(* IEC 61131-3 sources: Pirate/PLC/POU, 5 files *)

(* ---- EcrireSorties.st ---- *)
FUNCTION EcrireSorties : BOOL
// POU autonome extrait de FB_InterfacePIRATE (branche dev).
// A appeler APRES le calcul du simulateur.
// Reproduit uniquement les copies de variables GVL ; aucun mapping BFS ajoute.
// Appeler apres la simulation.
GVL_PIRATE.ST_THEGONNEC_AT2_Defaut_Auto_transfo_2 := GVL_PIRATE_Interne.S_ST_THEGONNEC_AT2_Defaut_Auto_transfo_2;
GVL_PIRATE.ST_THEGONNEC_SYSTEME_PC_SNCF_PA_Defaut_Controle_General := GVL_PIRATE_Interne.S_ST_THEGONNEC_SYSTEME_PC_SNCF_PA_Defaut_Controle_General;
GVL_PIRATE.ST_THEGONNEC_U_Cat__TT_2C_Etat_tension_voie_2 := GVL_PIRATE_Interne.S_ST_THEGONNEC_U_Cat__TT_2C_Etat_tension_voie_2;
GVL_PIRATE.ST_THEGONNEC_U_Cat__TT_3C_Etat_tension_voie_1 := GVL_PIRATE_Interne.S_ST_THEGONNEC_U_Cat__TT_3C_Etat_tension_voie_1;
GVL_PIRATE.ST_THEGONNEC_AT1_Defaut_Auto_transfo_1 := GVL_PIRATE_Interne.S_ST_THEGONNEC_AT1_Defaut_Auto_transfo_1;
GVL_PIRATE.BREST_SYSTEME_PC_SNCF_PA_Defaut_Controle_General := GVL_PIRATE_Interne.S_BREST_SYSTEME_PC_SNCF_PA_Defaut_Controle_General;
GVL_PIRATE.BREST_SA_Defaut_Chauffage_Commandes := GVL_PIRATE_Interne.S_BREST_SA_Defaut_Chauffage_Commandes;
GVL_PIRATE.BREST_U_Cat__TT_IA6_Etat_tension_voie := GVL_PIRATE_Interne.S_BREST_U_Cat__TT_IA6_Etat_tension_voie;
GVL_PIRATE.BREST_U_Cat__TT_IA1_Etat_tension_voie := GVL_PIRATE_Interne.S_BREST_U_Cat__TT_IA1_Etat_tension_voie;
GVL_PIRATE.BREST_U_Cat__TT_2C_Etat_tension_voie_2 := GVL_PIRATE_Interne.S_BREST_U_Cat__TT_2C_Etat_tension_voie_2;
GVL_PIRATE.PENCRAN_1_U_Feeder_TT_3F_Etat_tension_voie_1 := GVL_PIRATE_Interne.S_PENCRAN_1_U_Feeder_TT_3F_Etat_tension_voie_1;
GVL_PIRATE.PENCRAN_1_U_Feeder_TT_4F_Etat_tension_voie_2 := GVL_PIRATE_Interne.S_PENCRAN_1_U_Feeder_TT_4F_Etat_tension_voie_2;
GVL_PIRATE.PENCRAN_1_TT_Feeder_DL_Etat_tension := GVL_PIRATE_Interne.S_PENCRAN_1_TT_Feeder_DL_Etat_tension;
GVL_PIRATE.PENCRAN_1_U_Cat__TT_2C_Etat_tension_voie_2 := GVL_PIRATE_Interne.S_PENCRAN_1_U_Cat__TT_2C_Etat_tension_voie_2;
GVL_PIRATE.PENCRAN_1_U_Cat__TT_4C_Etat_tension_voie_2 := GVL_PIRATE_Interne.S_PENCRAN_1_U_Cat__TT_4C_Etat_tension_voie_2;
GVL_PIRATE.PENCRAN_1_U_Feeder_TT_1F_Etat_tension_voie_1 := GVL_PIRATE_Interne.S_PENCRAN_1_U_Feeder_TT_1F_Etat_tension_voie_1;
GVL_PIRATE.PENCRAN_1_U_Cat__TT_3C_Etat_tension_voie_1 := GVL_PIRATE_Interne.S_PENCRAN_1_U_Cat__TT_3C_Etat_tension_voie_1;
GVL_PIRATE.PENCRAN_1_U_Cat__TT_1C_Etat_tension_voie_1 := GVL_PIRATE_Interne.S_PENCRAN_1_U_Cat__TT_1C_Etat_tension_voie_1;
GVL_PIRATE.PENCRAN_1_TT_Cat__DB_Etat_tension := GVL_PIRATE_Interne.S_PENCRAN_1_TT_Cat__DB_Etat_tension;
GVL_PIRATE.PENCRAN_1_U_Feeder_TT_2F_Etat_tension_voie_2 := GVL_PIRATE_Interne.S_PENCRAN_1_U_Feeder_TT_2F_Etat_tension_voie_2;
GVL_PIRATE.PENCRAN_1_SYSTEME_PC_SNCF_PA_Defaut_Controle_General := GVL_PIRATE_Interne.S_PENCRAN_1_SYSTEME_PC_SNCF_PA_Defaut_Controle_General;
GVL_PIRATE.PENCRAN_1_TT_Cat__DL_Etat_tension := GVL_PIRATE_Interne.S_PENCRAN_1_TT_Cat__DL_Etat_tension;
GVL_PIRATE.PENCRAN_1_TT_Feeder_DB_Etat_tension := GVL_PIRATE_Interne.S_PENCRAN_1_TT_Feeder_DB_Etat_tension;
GVL_PIRATE.PENCRAN_1_GT2_Defaut_Alim__Protection__W_D_ := GVL_PIRATE_Interne.S_PENCRAN_1_GT2_Defaut_Alim__Protection__W_D_;
GVL_PIRATE.PENCRAN_1_DL__TSS__Defaut_Alim__Protection__W_D_ := GVL_PIRATE_Interne.S_PENCRAN_1_DL__TSS__Defaut_Alim__Protection__W_D_;
GVL_PIRATE.PENCRAN_1_GT1_Defaut_Alim__Protection__W_D_ := GVL_PIRATE_Interne.S_PENCRAN_1_GT1_Defaut_Alim__Protection__W_D_;
GVL_PIRATE.PENCRAN_1_GT1_Defaut_Transfo__Groupe_Traction := GVL_PIRATE_Interne.S_PENCRAN_1_GT1_Defaut_Transfo__Groupe_Traction;
GVL_PIRATE.PENCRAN_1_GT2_Defaut_Transfo__Groupe_Traction := GVL_PIRATE_Interne.S_PENCRAN_1_GT2_Defaut_Transfo__Groupe_Traction;
GVL_PIRATE.PENCRAN_1_DL__TSS__Defaut_SF6 := GVL_PIRATE_Interne.S_PENCRAN_1_DL__TSS__Defaut_SF6;
GVL_PIRATE.PENCRAN_1_SA_Defaut_Chargeur := GVL_PIRATE_Interne.S_PENCRAN_1_SA_Defaut_Chargeur;
GVL_PIRATE.PENCRAN_1_D2___25kV_Defaut_SF6_2eme_seuil := GVL_PIRATE_Interne.S_PENCRAN_1_D2___25kV_Defaut_SF6_2eme_seuil;
GVL_PIRATE.PENCRAN_1_DB__TSS__Defaut_Alim__Protection__W_D_ := GVL_PIRATE_Interne.S_PENCRAN_1_DB__TSS__Defaut_Alim__Protection__W_D_;
GVL_PIRATE.PENCRAN_1_Automate_Defaut_Relais_PROM := GVL_PIRATE_Interne.S_PENCRAN_1_Automate_Defaut_Relais_PROM;
GVL_PIRATE.PENCRAN_1_D2___25kV_Defaut_Commande_disjoncteur := GVL_PIRATE_Interne.S_PENCRAN_1_D2___25kV_Defaut_Commande_disjoncteur;
GVL_PIRATE.PENCRAN_1_Automate_Defaut_Reenclencheur := GVL_PIRATE_Interne.S_PENCRAN_1_Automate_Defaut_Reenclencheur;
GVL_PIRATE.PENCRAN_1_DB__TSS__Defaut_SF6 := GVL_PIRATE_Interne.S_PENCRAN_1_DB__TSS__Defaut_SF6;
GVL_PIRATE.LANDIVISIAU_AT2_Defaut_Auto_transfo_2 := GVL_PIRATE_Interne.S_LANDIVISIAU_AT2_Defaut_Auto_transfo_2;
GVL_PIRATE.LANDIVISIAU_U_Cat__TT_2C_Etat_tension_voie_2 := GVL_PIRATE_Interne.S_LANDIVISIAU_U_Cat__TT_2C_Etat_tension_voie_2;
GVL_PIRATE.LANDIVISIAU_AT1_Defaut_Auto_transfo_1 := GVL_PIRATE_Interne.S_LANDIVISIAU_AT1_Defaut_Auto_transfo_1;
GVL_PIRATE.LANDIVISIAU_SYSTEME_PC_SNCF_PA_Defaut_Controle_General := GVL_PIRATE_Interne.S_LANDIVISIAU_SYSTEME_PC_SNCF_PA_Defaut_Controle_General;
GVL_PIRATE.LANDIVISIAU_U_Cat__TT_3C_Etat_tension_voie_1 := GVL_PIRATE_Interne.S_LANDIVISIAU_U_Cat__TT_3C_Etat_tension_voie_1;
GVL_PIRATE.ST_MARC_U_Cat__TT_3C_Etat_tension_voie_1 := GVL_PIRATE_Interne.S_ST_MARC_U_Cat__TT_3C_Etat_tension_voie_1;
GVL_PIRATE.ST_MARC_SYSTEME_PC_SNCF_PA_Defaut_Controle_General := GVL_PIRATE_Interne.S_ST_MARC_SYSTEME_PC_SNCF_PA_Defaut_Controle_General;
GVL_PIRATE.ST_MARC_AT1_Defaut_Auto_transfo_1 := GVL_PIRATE_Interne.S_ST_MARC_AT1_Defaut_Auto_transfo_1;
GVL_PIRATE.ST_MARC_U_Cat__TT_2C_Etat_tension_voie_2 := GVL_PIRATE_Interne.S_ST_MARC_U_Cat__TT_2C_Etat_tension_voie_2;
GVL_PIRATE.ST_MARC_AT2_Defaut_Auto_transfo_2 := GVL_PIRATE_Interne.S_ST_MARC_AT2_Defaut_Auto_transfo_2;
GVL_PIRATE.LA_FOREST_AT_Defaut_Auto_transfo := GVL_PIRATE_Interne.S_LA_FOREST_AT_Defaut_Auto_transfo;
GVL_PIRATE.LA_FOREST_SYSTEME_PC_SNCF_PA_Defaut_Controle_General := GVL_PIRATE_Interne.S_LA_FOREST_SYSTEME_PC_SNCF_PA_Defaut_Controle_General;
GVL_PIRATE.KERIVIN_SYSTEME_PC_SNCF_PA_Defaut_Controle_General := GVL_PIRATE_Interne.S_KERIVIN_SYSTEME_PC_SNCF_PA_Defaut_Controle_General;
GVL_PIRATE.KERIVIN_U_Cat__TT_2C_Etat_tension_voie_2 := GVL_PIRATE_Interne.S_KERIVIN_U_Cat__TT_2C_Etat_tension_voie_2;
GVL_PIRATE.KERIVIN_AT2_Defaut_Auto_transfo_2 := GVL_PIRATE_Interne.S_KERIVIN_AT2_Defaut_Auto_transfo_2;
GVL_PIRATE.KERIVIN_AT1_Defaut_Auto_transfo_1 := GVL_PIRATE_Interne.S_KERIVIN_AT1_Defaut_Auto_transfo_1;
GVL_PIRATE.KERIVIN_U_Cat__TT_3C_Etat_tension_voie_1 := GVL_PIRATE_Interne.S_KERIVIN_U_Cat__TT_3C_Etat_tension_voie_1;
GVL_PIRATE.LANDERNEAU_SYSTEME_PC_SNCF_PA_Defaut_Controle_General := GVL_PIRATE_Interne.S_LANDERNEAU_SYSTEME_PC_SNCF_PA_Defaut_Controle_General;
GVL_PIRATE.MORLAIX_SYSTEME_PC_SNCF_PA_Defaut_Controle_General := GVL_PIRATE_Interne.S_MORLAIX_SYSTEME_PC_SNCF_PA_Defaut_Controle_General;
GVL_PIRATE.PLOUIGNEAU_U_Cat__TT_3C_Etat_tension_voie_1 := GVL_PIRATE_Interne.S_PLOUIGNEAU_U_Cat__TT_3C_Etat_tension_voie_1;
GVL_PIRATE.PLOUIGNEAU_U_Cat__TT_2C_Etat_tension_voie_2 := GVL_PIRATE_Interne.S_PLOUIGNEAU_U_Cat__TT_2C_Etat_tension_voie_2;
GVL_PIRATE.PLOUIGNEAU_AT1_Defaut_Auto_transfo_1 := GVL_PIRATE_Interne.S_PLOUIGNEAU_AT1_Defaut_Auto_transfo_1;
GVL_PIRATE.PLOUIGNEAU_U_Cat__TT_4C_Etat_tension_voie_2 := GVL_PIRATE_Interne.S_PLOUIGNEAU_U_Cat__TT_4C_Etat_tension_voie_2;
GVL_PIRATE.PLOUIGNEAU_AT2_Defaut_Auto_transfo_2 := GVL_PIRATE_Interne.S_PLOUIGNEAU_AT2_Defaut_Auto_transfo_2;
GVL_PIRATE.PLOUIGNEAU_SYSTEME_PC_SNCF_PA_Defaut_Controle_General := GVL_PIRATE_Interne.S_PLOUIGNEAU_SYSTEME_PC_SNCF_PA_Defaut_Controle_General;
GVL_PIRATE.PLOUNERIN_AT2_Defaut_Auto_transfo_2 := GVL_PIRATE_Interne.S_PLOUNERIN_AT2_Defaut_Auto_transfo_2;
GVL_PIRATE.PLOUNERIN_U_Cat__TT_3C_Etat_tension_voie_1 := GVL_PIRATE_Interne.S_PLOUNERIN_U_Cat__TT_3C_Etat_tension_voie_1;
EcrireSorties := TRUE;
END_FUNCTION

(* ---- LireEntrees.st ---- *)
FUNCTION LireEntrees : BOOL
// POU autonome extrait de FB_InterfacePIRATE (branche dev).
// A appeler AVANT le calcul du simulateur.
// Reproduit uniquement les copies de variables GVL ; aucun mapping BFS ajoute.
// Appeler avant la simulation.
GVL_PIRATE_Interne.E_ST_THEGONNEC_S20_30_Sect__de_pontage_V2 := GVL_PIRATE.ST_THEGONNEC_S20_30_Sect__de_pontage_V2;
GVL_PIRATE_Interne.E_ST_THEGONNEC_SYSTEME_PC_SNCF_PA_Douteux_vu_du_PC := GVL_PIRATE.ST_THEGONNEC_SYSTEME_PC_SNCF_PA_Douteux_vu_du_PC;
GVL_PIRATE_Interne.E_ST_THEGONNEC_IL2_Inter__de_ligne_2x25kv_V2 := GVL_PIRATE.ST_THEGONNEC_IL2_Inter__de_ligne_2x25kv_V2;
GVL_PIRATE_Interne.E_ST_THEGONNEC_IL4_Inter__de_ligne_2x25kv_V2 := GVL_PIRATE.ST_THEGONNEC_IL4_Inter__de_ligne_2x25kv_V2;
GVL_PIRATE_Interne.E_ST_THEGONNEC_SAT1___25kV_Sect__alimentation_auto_transfo1 := GVL_PIRATE.ST_THEGONNEC_SAT1___25kV_Sect__alimentation_auto_transfo1;
GVL_PIRATE_Interne.E_ST_THEGONNEC_SYSTEME_PC_SNCF_PA_Titulaire := GVL_PIRATE.ST_THEGONNEC_SYSTEME_PC_SNCF_PA_Titulaire;
GVL_PIRATE_Interne.E_ST_THEGONNEC_S21_31_Sect__de_pontage_V1 := GVL_PIRATE.ST_THEGONNEC_S21_31_Sect__de_pontage_V1;
GVL_PIRATE_Interne.E_ST_THEGONNEC_SYSTEME_PA_SNCF_PA_Perte_Date := GVL_PIRATE.ST_THEGONNEC_SYSTEME_PA_SNCF_PA_Perte_Date;
GVL_PIRATE_Interne.E_ST_THEGONNEC_IL3_Inter__de_ligne_2x25kv_V1 := GVL_PIRATE.ST_THEGONNEC_IL3_Inter__de_ligne_2x25kv_V1;
GVL_PIRATE_Interne.E_ST_THEGONNEC_SA_Manque_SA := GVL_PIRATE.ST_THEGONNEC_SA_Manque_SA;
GVL_PIRATE_Interne.E_ST_THEGONNEC_SYSTEME_PA_SNCF_PA_Carte_s__TS := GVL_PIRATE.ST_THEGONNEC_SYSTEME_PA_SNCF_PA_Carte_s__TS;
GVL_PIRATE_Interne.E_ST_THEGONNEC_IMP___25kV_Interrupteur_mise_en_parallele := GVL_PIRATE.ST_THEGONNEC_IMP___25kV_Interrupteur_mise_en_parallele;
GVL_PIRATE_Interne.E_ST_THEGONNEC_IL1_Inter__de_ligne_2x25kv_V1 := GVL_PIRATE.ST_THEGONNEC_IL1_Inter__de_ligne_2x25kv_V1;
GVL_PIRATE_Interne.E_ST_THEGONNEC_SYSTEME_PC_SNCF_PA_Liaison_PC______PA := GVL_PIRATE.ST_THEGONNEC_SYSTEME_PC_SNCF_PA_Liaison_PC______PA;
GVL_PIRATE_Interne.E_ST_THEGONNEC_SYSTEME_PC_SNCF_PA_Non_date := GVL_PIRATE.ST_THEGONNEC_SYSTEME_PC_SNCF_PA_Non_date;
GVL_PIRATE_Interne.E_ST_THEGONNEC_Contrile_Local_Commande_locale_individuelle := GVL_PIRATE.ST_THEGONNEC_Contrile_Local_Commande_locale_individuelle;
GVL_PIRATE_Interne.E_ST_THEGONNEC_FICTIF_Organe_Fictif := GVL_PIRATE.ST_THEGONNEC_FICTIF_Organe_Fictif;
GVL_PIRATE_Interne.E_ST_THEGONNEC_SAT2___25kV_Sect__alimentation_auto_transfo2 := GVL_PIRATE.ST_THEGONNEC_SAT2___25kV_Sect__alimentation_auto_transfo2;
GVL_PIRATE_Interne.E_ST_THEGONNEC_SYSTEME_PA_SNCF_PA_Perte_Information := GVL_PIRATE.ST_THEGONNEC_SYSTEME_PA_SNCF_PA_Perte_Information;
GVL_PIRATE_Interne.E_ST_THEGONNEC_SYSTEME_PA_SNCF_PA_Carte_s__TC := GVL_PIRATE.ST_THEGONNEC_SYSTEME_PA_SNCF_PA_Carte_s__TC;
GVL_PIRATE_Interne.E_BREST_SA_Manque_SA := GVL_PIRATE.BREST_SA_Manque_SA;
GVL_PIRATE_Interne.E_BREST_SYSTEME_PA_SNCF_PA_Carte_s__TS := GVL_PIRATE.BREST_SYSTEME_PA_SNCF_PA_Carte_s__TS;
GVL_PIRATE_Interne.E_BREST_Contrile_Local_Commande_locale_individuelle := GVL_PIRATE.BREST_Contrile_Local_Commande_locale_individuelle;
GVL_PIRATE_Interne.E_BREST_SYSTEME_PC_SNCF_PA_Non_date := GVL_PIRATE.BREST_SYSTEME_PC_SNCF_PA_Non_date;
GVL_PIRATE_Interne.E_BREST_SYSTEME_PA_SNCF_PA_Perte_Date := GVL_PIRATE.BREST_SYSTEME_PA_SNCF_PA_Perte_Date;
GVL_PIRATE_Interne.E_BREST_SYSTEME_PC_SNCF_PA_Liaison_PC______PA := GVL_PIRATE.BREST_SYSTEME_PC_SNCF_PA_Liaison_PC______PA;
GVL_PIRATE_Interne.E_BREST_SYSTEME_PA_SNCF_PA_Perte_Information := GVL_PIRATE.BREST_SYSTEME_PA_SNCF_PA_Perte_Information;
GVL_PIRATE_Interne.E_BREST_SYSTEME_PC_SNCF_PA_Titulaire := GVL_PIRATE.BREST_SYSTEME_PC_SNCF_PA_Titulaire;
GVL_PIRATE_Interne.E_BREST_IA6_Automatisme_Automat_Ouv_PLUS_Bloc_Debloc_IA__Ouv_ := GVL_PIRATE.BREST_IA6_Automatisme_Automat_Ouv_PLUS_Bloc_Debloc_IA__Ouv_;
GVL_PIRATE_Interne.E_BREST_IL2_Inter__de_ligne_25kv_V2 := GVL_PIRATE.BREST_IL2_Inter__de_ligne_25kv_V2;
GVL_PIRATE_Interne.E_BREST_IA1_Automatisme_Automat_Ouv_PLUS_Bloc_Debloc_IA__Ouv_ := GVL_PIRATE.BREST_IA1_Automatisme_Automat_Ouv_PLUS_Bloc_Debloc_IA__Ouv_;
GVL_PIRATE_Interne.E_BREST_IA6_Interrupteur_d_Alimentation__IA_ := GVL_PIRATE.BREST_IA6_Interrupteur_d_Alimentation__IA_;
GVL_PIRATE_Interne.E_BREST_IL1_Inter__de_ligne_25kv_V1 := GVL_PIRATE.BREST_IL1_Inter__de_ligne_25kv_V1;
GVL_PIRATE_Interne.E_BREST_SYSTEME_PC_SNCF_PA_Douteux_vu_du_PC := GVL_PIRATE.BREST_SYSTEME_PC_SNCF_PA_Douteux_vu_du_PC;
GVL_PIRATE_Interne.E_BREST_IA1_Interrupteur_d_Alimentation__IA_ := GVL_PIRATE.BREST_IA1_Interrupteur_d_Alimentation__IA_;
GVL_PIRATE_Interne.E_BREST_SYSTEME_PA_SNCF_PA_Carte_s__TC := GVL_PIRATE.BREST_SYSTEME_PA_SNCF_PA_Carte_s__TC;
GVL_PIRATE_Interne.E_BREST_FICTIF_Organe_Fictif := GVL_PIRATE.BREST_FICTIF_Organe_Fictif;
GVL_PIRATE_Interne.E_PENCRAN_1_SYSTEME_PC_SNCF_PA_Douteux_vu_du_PC := GVL_PIRATE.PENCRAN_1_SYSTEME_PC_SNCF_PA_Douteux_vu_du_PC;
GVL_PIRATE_Interne.E_PENCRAN_1_SYSTEME_PA_SNCF_PA_Perte_Date := GVL_PIRATE.PENCRAN_1_SYSTEME_PA_SNCF_PA_Perte_Date;
GVL_PIRATE_Interne.E_PENCRAN_1_SYSTEME_PC_SNCF_PA_Non_date := GVL_PIRATE.PENCRAN_1_SYSTEME_PC_SNCF_PA_Non_date;
GVL_PIRATE_Interne.E_PENCRAN_1_UHT_1_Absence_tension_ligne_HT := GVL_PIRATE.PENCRAN_1_UHT_1_Absence_tension_ligne_HT;
GVL_PIRATE_Interne.E_PENCRAN_1_SYSTEME_PC_SNCF_PA_Liaison_PC______PA := GVL_PIRATE.PENCRAN_1_SYSTEME_PC_SNCF_PA_Liaison_PC______PA;
GVL_PIRATE_Interne.E_PENCRAN_1_SYSTEME_PA_SNCF_PA_Perte_Information := GVL_PIRATE.PENCRAN_1_SYSTEME_PA_SNCF_PA_Perte_Information;
GVL_PIRATE_Interne.E_PENCRAN_1_UHT_1_Fusion_fusible_s_ := GVL_PIRATE.PENCRAN_1_UHT_1_Fusion_fusible_s_;
GVL_PIRATE_Interne.E_PENCRAN_1_SYSTEME_PC_SNCF_PA_Titulaire := GVL_PIRATE.PENCRAN_1_SYSTEME_PC_SNCF_PA_Titulaire;
GVL_PIRATE_Interne.E_PENCRAN_1_UHT_2_Absence_tension_ligne_HT := GVL_PIRATE.PENCRAN_1_UHT_2_Absence_tension_ligne_HT;
GVL_PIRATE_Interne.E_PENCRAN_1_UHT_2_Fusion_fusible_s_ := GVL_PIRATE.PENCRAN_1_UHT_2_Fusion_fusible_s_;
GVL_PIRATE_Interne.E_PENCRAN_1_SLB1_Sect__de_barre_de_ligne_25Kv := GVL_PIRATE.PENCRAN_1_SLB1_Sect__de_barre_de_ligne_25Kv;
GVL_PIRATE_Interne.E_PENCRAN_1_DL_Disj_depart_2x25kV_Le_Mans := GVL_PIRATE.PENCRAN_1_DL_Disj_depart_2x25kV_Le_Mans;
GVL_PIRATE_Interne.E_PENCRAN_1_S11___63kV_Sect__de_ligne_Haute_Tension := GVL_PIRATE.PENCRAN_1_S11___63kV_Sect__de_ligne_Haute_Tension;
GVL_PIRATE_Interne.E_PENCRAN_1_SA_Manque_SA2 := GVL_PIRATE.PENCRAN_1_SA_Manque_SA2;
GVL_PIRATE_Interne.E_PENCRAN_1_IS1_Inter__de_S_Station_2x25Kv_V1 := GVL_PIRATE.PENCRAN_1_IS1_Inter__de_S_Station_2x25Kv_V1;
GVL_PIRATE_Interne.E_PENCRAN_1_SRB1___25kV_Sect__a_rupture_brusque_GT1 := GVL_PIRATE.PENCRAN_1_SRB1___25kV_Sect__a_rupture_brusque_GT1;
GVL_PIRATE_Interne.E_PENCRAN_1_SYSTEME_PA_SNCF_PA_Carte_s__TS := GVL_PIRATE.PENCRAN_1_SYSTEME_PA_SNCF_PA_Carte_s__TS;
GVL_PIRATE_Interne.E_PENCRAN_1_SA_Manque_SA1 := GVL_PIRATE.PENCRAN_1_SA_Manque_SA1;
GVL_PIRATE_Interne.E_PENCRAN_1_SA_Manque_48V_ := GVL_PIRATE.PENCRAN_1_SA_Manque_48V_;
GVL_PIRATE_Interne.E_PENCRAN_1_SYSTEME_PA_SNCF_PA_Carte_s__TC := GVL_PIRATE.PENCRAN_1_SYSTEME_PA_SNCF_PA_Carte_s__TC;
GVL_PIRATE_Interne.E_PENCRAN_1_P1_Sect__de_pontage_V1 := GVL_PIRATE.PENCRAN_1_P1_Sect__de_pontage_V1;
GVL_PIRATE_Interne.E_PENCRAN_1_SB1___25kV_Sect__de_section_de_barre_25Kv := GVL_PIRATE.PENCRAN_1_SB1___25kV_Sect__de_section_de_barre_25Kv;
GVL_PIRATE_Interne.E_PENCRAN_1_SBP1___63kV_Sect__de_section_de_barre_HT := GVL_PIRATE.PENCRAN_1_SBP1___63kV_Sect__de_section_de_barre_HT;
GVL_PIRATE_Interne.E_PENCRAN_1_IS3_Inter__de_S_Station_25Kv_V1 := GVL_PIRATE.PENCRAN_1_IS3_Inter__de_S_Station_25Kv_V1;
GVL_PIRATE_Interne.E_PENCRAN_1_P2_Sect__de_pontage_V2 := GVL_PIRATE.PENCRAN_1_P2_Sect__de_pontage_V2;
GVL_PIRATE_Interne.E_PENCRAN_1_IS2_Inter__de_S_Station_2x25Kv_V2 := GVL_PIRATE.PENCRAN_1_IS2_Inter__de_S_Station_2x25Kv_V2;
GVL_PIRATE_Interne.E_PENCRAN_1_S21___63kV_Sect__de_ligne_Haute_Tension := GVL_PIRATE.PENCRAN_1_S21___63kV_Sect__de_ligne_Haute_Tension;
GVL_PIRATE_Interne.E_PENCRAN_1_IS4_Inter__de_S_Station_2x25Kv_V2 := GVL_PIRATE.PENCRAN_1_IS4_Inter__de_S_Station_2x25Kv_V2;
GVL_PIRATE_Interne.E_PENCRAN_1_SRB2___25kV_Sect__a_rupture_brusque_GT2 := GVL_PIRATE.PENCRAN_1_SRB2___25kV_Sect__a_rupture_brusque_GT2;
GVL_PIRATE_Interne.E_PENCRAN_1_D2___63kV_Disjoncteur_Groupe_Traction_2 := GVL_PIRATE.PENCRAN_1_D2___63kV_Disjoncteur_Groupe_Traction_2;
GVL_PIRATE_Interne.E_PENCRAN_1_DB_Disj_depart_2x25kV_Brest := GVL_PIRATE.PENCRAN_1_DB_Disj_depart_2x25kV_Brest;
GVL_PIRATE_Interne.E_PENCRAN_1_D2___25kV_Alarme_SF6_1er_seuil := GVL_PIRATE.PENCRAN_1_D2___25kV_Alarme_SF6_1er_seuil;
GVL_PIRATE_Interne.E_PENCRAN_1_Automate_Relais_PROM__TC_ := GVL_PIRATE.PENCRAN_1_Automate_Relais_PROM__TC_;
GVL_PIRATE_Interne.E_PENCRAN_1_Contrile_Local_Commande_Locale := GVL_PIRATE.PENCRAN_1_Contrile_Local_Commande_Locale;
GVL_PIRATE_Interne.E_PENCRAN_1_D1___63kV_Disjoncteur_Groupe_Traction_1 := GVL_PIRATE.PENCRAN_1_D1___63kV_Disjoncteur_Groupe_Traction_1;
GVL_PIRATE_Interne.E_PENCRAN_1_VF_Veille_Franchissement__TC_ := GVL_PIRATE.PENCRAN_1_VF_Veille_Franchissement__TC_;
GVL_PIRATE_Interne.E_PENCRAN_1_FICTIF_Organe_Fictif := GVL_PIRATE.PENCRAN_1_FICTIF_Organe_Fictif;
GVL_PIRATE_Interne.E_PENCRAN_1_D2___25kV_Disjoncteur_Groupe_Traction_2 := GVL_PIRATE.PENCRAN_1_D2___25kV_Disjoncteur_Groupe_Traction_2;
GVL_PIRATE_Interne.E_LANDIVISIAU_SYSTEME_PA_SNCF_PA_Perte_Date := GVL_PIRATE.LANDIVISIAU_SYSTEME_PA_SNCF_PA_Perte_Date;
GVL_PIRATE_Interne.E_LANDIVISIAU_S30_40_Sect__de_pontage_V2 := GVL_PIRATE.LANDIVISIAU_S30_40_Sect__de_pontage_V2;
GVL_PIRATE_Interne.E_LANDIVISIAU_SYSTEME_PC_SNCF_PA_Non_date := GVL_PIRATE.LANDIVISIAU_SYSTEME_PC_SNCF_PA_Non_date;
GVL_PIRATE_Interne.E_LANDIVISIAU_S31_41_Sect__de_pontage_V1 := GVL_PIRATE.LANDIVISIAU_S31_41_Sect__de_pontage_V1;
GVL_PIRATE_Interne.E_LANDIVISIAU_IL1_Inter__de_ligne_2x25kv_V1 := GVL_PIRATE.LANDIVISIAU_IL1_Inter__de_ligne_2x25kv_V1;
GVL_PIRATE_Interne.E_LANDIVISIAU_SYSTEME_PC_SNCF_PA_Douteux_vu_du_PC := GVL_PIRATE.LANDIVISIAU_SYSTEME_PC_SNCF_PA_Douteux_vu_du_PC;
GVL_PIRATE_Interne.E_LANDIVISIAU_SYSTEME_PA_SNCF_PA_Carte_s__TS := GVL_PIRATE.LANDIVISIAU_SYSTEME_PA_SNCF_PA_Carte_s__TS;
GVL_PIRATE_Interne.E_LANDIVISIAU_IL3_Inter__de_ligne_2x25kv_V1 := GVL_PIRATE.LANDIVISIAU_IL3_Inter__de_ligne_2x25kv_V1;
GVL_PIRATE_Interne.E_LANDIVISIAU_SA_Manque_SA := GVL_PIRATE.LANDIVISIAU_SA_Manque_SA;
GVL_PIRATE_Interne.E_LANDIVISIAU_SYSTEME_PC_SNCF_PA_Liaison_PC______PA := GVL_PIRATE.LANDIVISIAU_SYSTEME_PC_SNCF_PA_Liaison_PC______PA;
GVL_PIRATE_Interne.E_LANDIVISIAU_IL2_Inter__de_ligne_2x25kv_V2 := GVL_PIRATE.LANDIVISIAU_IL2_Inter__de_ligne_2x25kv_V2;
GVL_PIRATE_Interne.E_LANDIVISIAU_IMP___25kV_Interrupteur_mise_en_parallele := GVL_PIRATE.LANDIVISIAU_IMP___25kV_Interrupteur_mise_en_parallele;
GVL_PIRATE_Interne.E_LANDIVISIAU_SAT1___25kV_Sect__alimentation_auto_transfo1 := GVL_PIRATE.LANDIVISIAU_SAT1___25kV_Sect__alimentation_auto_transfo1;
GVL_PIRATE_Interne.E_LANDIVISIAU_SYSTEME_PC_SNCF_PA_Titulaire := GVL_PIRATE.LANDIVISIAU_SYSTEME_PC_SNCF_PA_Titulaire;
GVL_PIRATE_Interne.E_LANDIVISIAU_IL4_Inter__de_ligne_2x25kv_V2 := GVL_PIRATE.LANDIVISIAU_IL4_Inter__de_ligne_2x25kv_V2;
GVL_PIRATE_Interne.E_LANDIVISIAU_SYSTEME_PA_SNCF_PA_Perte_Information := GVL_PIRATE.LANDIVISIAU_SYSTEME_PA_SNCF_PA_Perte_Information;
GVL_PIRATE_Interne.E_LANDIVISIAU_SYSTEME_PA_SNCF_PA_Carte_s__TC := GVL_PIRATE.LANDIVISIAU_SYSTEME_PA_SNCF_PA_Carte_s__TC;
GVL_PIRATE_Interne.E_LANDIVISIAU_Contrile_Local_Commande_locale_individuelle := GVL_PIRATE.LANDIVISIAU_Contrile_Local_Commande_locale_individuelle;
GVL_PIRATE_Interne.E_LANDIVISIAU_SAT2___25kV_Sect__alimentation_auto_transfo2 := GVL_PIRATE.LANDIVISIAU_SAT2___25kV_Sect__alimentation_auto_transfo2;
GVL_PIRATE_Interne.E_LANDIVISIAU_FICTIF_Organe_Fictif := GVL_PIRATE.LANDIVISIAU_FICTIF_Organe_Fictif;
GVL_PIRATE_Interne.E_ST_MARC_S4_10_Sect__de_pontage_V2 := GVL_PIRATE.ST_MARC_S4_10_Sect__de_pontage_V2;
GVL_PIRATE_Interne.E_ST_MARC_SYSTEME_PA_SNCF_PA_Perte_Information := GVL_PIRATE.ST_MARC_SYSTEME_PA_SNCF_PA_Perte_Information;
GVL_PIRATE_Interne.E_ST_MARC_IA3_Interrupteur_d_Alimentation__IA_ := GVL_PIRATE.ST_MARC_IA3_Interrupteur_d_Alimentation__IA_;
GVL_PIRATE_Interne.E_ST_MARC_SA_Manque_SA_Satellite_2 := GVL_PIRATE.ST_MARC_SA_Manque_SA_Satellite_2;
GVL_PIRATE_Interne.E_ST_MARC_IL2_Inter__de_ligne_2x25kv_V2 := GVL_PIRATE.ST_MARC_IL2_Inter__de_ligne_2x25kv_V2;
GVL_PIRATE_Interne.E_ST_MARC_IMP___25kV_Interrupteur_mise_en_parallele := GVL_PIRATE.ST_MARC_IMP___25kV_Interrupteur_mise_en_parallele;
GVL_PIRATE_Interne.E_ST_MARC_SYSTEME_PC_SNCF_PA_Non_date := GVL_PIRATE.ST_MARC_SYSTEME_PC_SNCF_PA_Non_date;
GVL_PIRATE_Interne.E_ST_MARC_SYSTEME_PA_SNCF_PA_Carte_s__TS := GVL_PIRATE.ST_MARC_SYSTEME_PA_SNCF_PA_Carte_s__TS;
GVL_PIRATE_Interne.E_ST_MARC_I5_Interrupteur_2x25kV_V1 := GVL_PIRATE.ST_MARC_I5_Interrupteur_2x25kV_V1;
GVL_PIRATE_Interne.E_ST_MARC_SA_Manque_SA := GVL_PIRATE.ST_MARC_SA_Manque_SA;
GVL_PIRATE_Interne.E_ST_MARC_IL4_Inter__de_ligne_25kv_V2 := GVL_PIRATE.ST_MARC_IL4_Inter__de_ligne_25kv_V2;
GVL_PIRATE_Interne.E_ST_MARC_SA_Manque_SA_Satellite_1 := GVL_PIRATE.ST_MARC_SA_Manque_SA_Satellite_1;
GVL_PIRATE_Interne.E_ST_MARC_IL1_Inter__de_ligne_2x25kv_V1 := GVL_PIRATE.ST_MARC_IL1_Inter__de_ligne_2x25kv_V1;
GVL_PIRATE_Interne.E_ST_MARC_SYSTEME_PA_SNCF_PA_Perte_Date := GVL_PIRATE.ST_MARC_SYSTEME_PA_SNCF_PA_Perte_Date;
GVL_PIRATE_Interne.E_ST_MARC_IL3_Inter__de_ligne_25kv_V1 := GVL_PIRATE.ST_MARC_IL3_Inter__de_ligne_25kv_V1;
GVL_PIRATE_Interne.E_ST_MARC_SYSTEME_PC_SNCF_PA_Douteux_vu_du_PC := GVL_PIRATE.ST_MARC_SYSTEME_PC_SNCF_PA_Douteux_vu_du_PC;
GVL_PIRATE_Interne.E_ST_MARC_SAT2___25kV_Sect__alimentation_auto_transfo2 := GVL_PIRATE.ST_MARC_SAT2___25kV_Sect__alimentation_auto_transfo2;
GVL_PIRATE_Interne.E_ST_MARC_S5_11_Sect__de_pontage_V1 := GVL_PIRATE.ST_MARC_S5_11_Sect__de_pontage_V1;
GVL_PIRATE_Interne.E_ST_MARC_IA3_Automatisme_Automat_Ouv_PLUS_Bloc_Debloc_IA__Ouv_ := GVL_PIRATE.ST_MARC_IA3_Automatisme_Automat_Ouv_PLUS_Bloc_Debloc_IA__Ouv_;
GVL_PIRATE_Interne.E_ST_MARC_SYSTEME_PC_SNCF_PA_Liaison_PC______PA := GVL_PIRATE.ST_MARC_SYSTEME_PC_SNCF_PA_Liaison_PC______PA;
GVL_PIRATE_Interne.E_ST_MARC_Contrile_Local_Commande_locale_individuelle := GVL_PIRATE.ST_MARC_Contrile_Local_Commande_locale_individuelle;
GVL_PIRATE_Interne.E_ST_MARC_SAT1___25kV_Sect__alimentation_auto_transfo1 := GVL_PIRATE.ST_MARC_SAT1___25kV_Sect__alimentation_auto_transfo1;
GVL_PIRATE_Interne.E_ST_MARC_SYSTEME_PC_SNCF_PA_Titulaire := GVL_PIRATE.ST_MARC_SYSTEME_PC_SNCF_PA_Titulaire;
GVL_PIRATE_Interne.E_ST_MARC_SYSTEME_PA_SNCF_PA_Carte_s__TC := GVL_PIRATE.ST_MARC_SYSTEME_PA_SNCF_PA_Carte_s__TC;
GVL_PIRATE_Interne.E_ST_MARC_FICTIF_Organe_Fictif := GVL_PIRATE.ST_MARC_FICTIF_Organe_Fictif;
GVL_PIRATE_Interne.E_LA_FOREST_SYSTEME_PA_SNCF_PA_Perte_Information := GVL_PIRATE.LA_FOREST_SYSTEME_PA_SNCF_PA_Perte_Information;
GVL_PIRATE_Interne.E_LA_FOREST_SYSTEME_PA_SNCF_PA_Carte_s__TS := GVL_PIRATE.LA_FOREST_SYSTEME_PA_SNCF_PA_Carte_s__TS;
GVL_PIRATE_Interne.E_LA_FOREST_SYSTEME_PA_SNCF_PA_Carte_s__TC := GVL_PIRATE.LA_FOREST_SYSTEME_PA_SNCF_PA_Carte_s__TC;
GVL_PIRATE_Interne.E_LA_FOREST_SYSTEME_PC_SNCF_PA_Liaison_PC______PA := GVL_PIRATE.LA_FOREST_SYSTEME_PC_SNCF_PA_Liaison_PC______PA;
GVL_PIRATE_Interne.E_LA_FOREST_SYSTEME_PA_SNCF_PA_Perte_Date := GVL_PIRATE.LA_FOREST_SYSTEME_PA_SNCF_PA_Perte_Date;
GVL_PIRATE_Interne.E_LA_FOREST_IMP2_Inter__mise_parallele_2x25kv_V2 := GVL_PIRATE.LA_FOREST_IMP2_Inter__mise_parallele_2x25kv_V2;
GVL_PIRATE_Interne.E_LA_FOREST_SYSTEME_PC_SNCF_PA_Titulaire := GVL_PIRATE.LA_FOREST_SYSTEME_PC_SNCF_PA_Titulaire;
GVL_PIRATE_Interne.E_LA_FOREST_SYSTEME_PC_SNCF_PA_Non_date := GVL_PIRATE.LA_FOREST_SYSTEME_PC_SNCF_PA_Non_date;
GVL_PIRATE_Interne.E_LA_FOREST_IMP1_Inter__mise_parallele_2x25kv_V1 := GVL_PIRATE.LA_FOREST_IMP1_Inter__mise_parallele_2x25kv_V1;
GVL_PIRATE_Interne.E_LA_FOREST_Contrile_Local_Commande_locale_individuelle := GVL_PIRATE.LA_FOREST_Contrile_Local_Commande_locale_individuelle;
GVL_PIRATE_Interne.E_LA_FOREST_SAT___25kV_Sect__alimentation_auto_transfo := GVL_PIRATE.LA_FOREST_SAT___25kV_Sect__alimentation_auto_transfo;
GVL_PIRATE_Interne.E_LA_FOREST_SA_Manque_SA := GVL_PIRATE.LA_FOREST_SA_Manque_SA;
GVL_PIRATE_Interne.E_LA_FOREST_SYSTEME_PC_SNCF_PA_Douteux_vu_du_PC := GVL_PIRATE.LA_FOREST_SYSTEME_PC_SNCF_PA_Douteux_vu_du_PC;
GVL_PIRATE_Interne.E_LA_FOREST_FICTIF_Organe_Fictif := GVL_PIRATE.LA_FOREST_FICTIF_Organe_Fictif;
GVL_PIRATE_Interne.E_KERIVIN_SAT1___25kV_Sect__alimentation_auto_transfo1 := GVL_PIRATE.KERIVIN_SAT1___25kV_Sect__alimentation_auto_transfo1;
GVL_PIRATE_Interne.E_KERIVIN_SYSTEME_PC_SNCF_PA_Douteux_vu_du_PC := GVL_PIRATE.KERIVIN_SYSTEME_PC_SNCF_PA_Douteux_vu_du_PC;
GVL_PIRATE_Interne.E_KERIVIN_SYSTEME_PC_SNCF_PA_Titulaire := GVL_PIRATE.KERIVIN_SYSTEME_PC_SNCF_PA_Titulaire;
GVL_PIRATE_Interne.E_KERIVIN_IL1_Inter__de_ligne_2x25kv_V1 := GVL_PIRATE.KERIVIN_IL1_Inter__de_ligne_2x25kv_V1;
GVL_PIRATE_Interne.E_KERIVIN_S18_20_Sect__de_pontage_V2 := GVL_PIRATE.KERIVIN_S18_20_Sect__de_pontage_V2;
GVL_PIRATE_Interne.E_KERIVIN_SYSTEME_PC_SNCF_PA_Liaison_PC______PA := GVL_PIRATE.KERIVIN_SYSTEME_PC_SNCF_PA_Liaison_PC______PA;
GVL_PIRATE_Interne.E_KERIVIN_SYSTEME_PA_SNCF_PA_Carte_s__TC := GVL_PIRATE.KERIVIN_SYSTEME_PA_SNCF_PA_Carte_s__TC;
GVL_PIRATE_Interne.E_KERIVIN_IL3_Inter__de_ligne_2x25kv_V1 := GVL_PIRATE.KERIVIN_IL3_Inter__de_ligne_2x25kv_V1;
GVL_PIRATE_Interne.E_KERIVIN_SA_Manque_SA := GVL_PIRATE.KERIVIN_SA_Manque_SA;
GVL_PIRATE_Interne.E_KERIVIN_SYSTEME_PA_SNCF_PA_Perte_Date := GVL_PIRATE.KERIVIN_SYSTEME_PA_SNCF_PA_Perte_Date;
GVL_PIRATE_Interne.E_KERIVIN_IMP___25kV_Interrupteur_mise_en_parallele := GVL_PIRATE.KERIVIN_IMP___25kV_Interrupteur_mise_en_parallele;
GVL_PIRATE_Interne.E_KERIVIN_SYSTEME_PA_SNCF_PA_Carte_s__TS := GVL_PIRATE.KERIVIN_SYSTEME_PA_SNCF_PA_Carte_s__TS;
GVL_PIRATE_Interne.E_KERIVIN_SYSTEME_PA_SNCF_PA_Perte_Information := GVL_PIRATE.KERIVIN_SYSTEME_PA_SNCF_PA_Perte_Information;
GVL_PIRATE_Interne.E_KERIVIN_IL2_Inter__de_ligne_2x25kv_V2 := GVL_PIRATE.KERIVIN_IL2_Inter__de_ligne_2x25kv_V2;
GVL_PIRATE_Interne.E_KERIVIN_SAT2___25kV_Sect__alimentation_auto_transfo2 := GVL_PIRATE.KERIVIN_SAT2___25kV_Sect__alimentation_auto_transfo2;
GVL_PIRATE_Interne.E_KERIVIN_SYSTEME_PC_SNCF_PA_Non_date := GVL_PIRATE.KERIVIN_SYSTEME_PC_SNCF_PA_Non_date;
GVL_PIRATE_Interne.E_KERIVIN_Contrile_Local_Commande_locale_individuelle := GVL_PIRATE.KERIVIN_Contrile_Local_Commande_locale_individuelle;
GVL_PIRATE_Interne.E_KERIVIN_S13_21_Sect__de_pontage_V1 := GVL_PIRATE.KERIVIN_S13_21_Sect__de_pontage_V1;
GVL_PIRATE_Interne.E_KERIVIN_IL4_Inter__de_ligne_2x25kv_V2 := GVL_PIRATE.KERIVIN_IL4_Inter__de_ligne_2x25kv_V2;
GVL_PIRATE_Interne.E_KERIVIN_FICTIF_Organe_Fictif := GVL_PIRATE.KERIVIN_FICTIF_Organe_Fictif;
GVL_PIRATE_Interne.E_LANDERNEAU_SYSTEME_PA_SNCF_PA_Perte_Date := GVL_PIRATE.LANDERNEAU_SYSTEME_PA_SNCF_PA_Perte_Date;
GVL_PIRATE_Interne.E_LANDERNEAU_SA_Manque_SA := GVL_PIRATE.LANDERNEAU_SA_Manque_SA;
GVL_PIRATE_Interne.E_LANDERNEAU_SYSTEME_PA_SNCF_PA_Carte_s__TS := GVL_PIRATE.LANDERNEAU_SYSTEME_PA_SNCF_PA_Carte_s__TS;
GVL_PIRATE_Interne.E_LANDERNEAU_I4_Interrupteur_2x25kV_V2 := GVL_PIRATE.LANDERNEAU_I4_Interrupteur_2x25kV_V2;
GVL_PIRATE_Interne.E_LANDERNEAU_I3_Interrupteur_2x25kV_V1 := GVL_PIRATE.LANDERNEAU_I3_Interrupteur_2x25kV_V1;
GVL_PIRATE_Interne.E_LANDERNEAU_SYSTEME_PA_SNCF_PA_Carte_s__TC := GVL_PIRATE.LANDERNEAU_SYSTEME_PA_SNCF_PA_Carte_s__TC;
GVL_PIRATE_Interne.E_LANDERNEAU_SYSTEME_PA_SNCF_PA_Perte_Information := GVL_PIRATE.LANDERNEAU_SYSTEME_PA_SNCF_PA_Perte_Information;
GVL_PIRATE_Interne.E_LANDERNEAU_SYSTEME_PC_SNCF_PA_Douteux_vu_du_PC := GVL_PIRATE.LANDERNEAU_SYSTEME_PC_SNCF_PA_Douteux_vu_du_PC;
GVL_PIRATE_Interne.E_LANDERNEAU_SYSTEME_PC_SNCF_PA_Liaison_PC______PA := GVL_PIRATE.LANDERNEAU_SYSTEME_PC_SNCF_PA_Liaison_PC______PA;
GVL_PIRATE_Interne.E_LANDERNEAU_SYSTEME_PC_SNCF_PA_Non_date := GVL_PIRATE.LANDERNEAU_SYSTEME_PC_SNCF_PA_Non_date;
GVL_PIRATE_Interne.E_LANDERNEAU_SYSTEME_PC_SNCF_PA_Titulaire := GVL_PIRATE.LANDERNEAU_SYSTEME_PC_SNCF_PA_Titulaire;
GVL_PIRATE_Interne.E_LANDERNEAU_Contrile_Local_Commande_locale_individuelle := GVL_PIRATE.LANDERNEAU_Contrile_Local_Commande_locale_individuelle;
GVL_PIRATE_Interne.E_LANDERNEAU_FICTIF_Organe_Fictif := GVL_PIRATE.LANDERNEAU_FICTIF_Organe_Fictif;
GVL_PIRATE_Interne.E_MORLAIX_SYSTEME_PA_SNCF_PA_Carte_s__TC := GVL_PIRATE.MORLAIX_SYSTEME_PA_SNCF_PA_Carte_s__TC;
GVL_PIRATE_Interne.E_MORLAIX_SA_Manque_SA := GVL_PIRATE.MORLAIX_SA_Manque_SA;
GVL_PIRATE_Interne.E_MORLAIX_SYSTEME_PC_SNCF_PA_Douteux_vu_du_PC := GVL_PIRATE.MORLAIX_SYSTEME_PC_SNCF_PA_Douteux_vu_du_PC;
GVL_PIRATE_Interne.E_MORLAIX_SA_Manque_SA_Satellite_1 := GVL_PIRATE.MORLAIX_SA_Manque_SA_Satellite_1;
GVL_PIRATE_Interne.E_MORLAIX_SYSTEME_PA_SNCF_PA_Perte_Date := GVL_PIRATE.MORLAIX_SYSTEME_PA_SNCF_PA_Perte_Date;
GVL_PIRATE_Interne.E_MORLAIX_SA_Manque_SA_Satellite_2 := GVL_PIRATE.MORLAIX_SA_Manque_SA_Satellite_2;
GVL_PIRATE_Interne.E_MORLAIX_Contrile_Local_Commande_locale_individuelle := GVL_PIRATE.MORLAIX_Contrile_Local_Commande_locale_individuelle;
GVL_PIRATE_Interne.E_MORLAIX_SYSTEME_PC_SNCF_PA_Liaison_PC______PA := GVL_PIRATE.MORLAIX_SYSTEME_PC_SNCF_PA_Liaison_PC______PA;
GVL_PIRATE_Interne.E_MORLAIX_I14_Interrupteur_2x25kV_V2 := GVL_PIRATE.MORLAIX_I14_Interrupteur_2x25kV_V2;
GVL_PIRATE_Interne.E_MORLAIX_I16_Inter__de_ligne_2x25kv_V2 := GVL_PIRATE.MORLAIX_I16_Inter__de_ligne_2x25kv_V2;
GVL_PIRATE_Interne.E_MORLAIX_I13_Interrupteur_2x25kV_V1 := GVL_PIRATE.MORLAIX_I13_Interrupteur_2x25kV_V1;
GVL_PIRATE_Interne.E_MORLAIX_I18_Interrupteur_2x25kV_V2 := GVL_PIRATE.MORLAIX_I18_Interrupteur_2x25kV_V2;
GVL_PIRATE_Interne.E_MORLAIX_SYSTEME_PA_SNCF_PA_Perte_Information := GVL_PIRATE.MORLAIX_SYSTEME_PA_SNCF_PA_Perte_Information;
GVL_PIRATE_Interne.E_MORLAIX_SYSTEME_PC_SNCF_PA_Non_date := GVL_PIRATE.MORLAIX_SYSTEME_PC_SNCF_PA_Non_date;
GVL_PIRATE_Interne.E_MORLAIX_SYSTEME_PA_SNCF_PA_Carte_s__TS := GVL_PIRATE.MORLAIX_SYSTEME_PA_SNCF_PA_Carte_s__TS;
GVL_PIRATE_Interne.E_MORLAIX_SYSTEME_PC_SNCF_PA_Titulaire := GVL_PIRATE.MORLAIX_SYSTEME_PC_SNCF_PA_Titulaire;
GVL_PIRATE_Interne.E_MORLAIX_FICTIF_Organe_Fictif := GVL_PIRATE.MORLAIX_FICTIF_Organe_Fictif;
GVL_PIRATE_Interne.E_PLOUIGNEAU_IL3_Inter__de_ligne_2x25kv_V1 := GVL_PIRATE.PLOUIGNEAU_IL3_Inter__de_ligne_2x25kv_V1;
GVL_PIRATE_Interne.E_PLOUIGNEAU_IMP___25kV_Interrupteur_mise_en_parallele := GVL_PIRATE.PLOUIGNEAU_IMP___25kV_Interrupteur_mise_en_parallele;
GVL_PIRATE_Interne.E_PLOUIGNEAU_SYSTEME_PA_SNCF_PA_Carte_s__TS := GVL_PIRATE.PLOUIGNEAU_SYSTEME_PA_SNCF_PA_Carte_s__TS;
GVL_PIRATE_Interne.E_PLOUIGNEAU_SYSTEME_PC_SNCF_PA_Liaison_PC______PA := GVL_PIRATE.PLOUIGNEAU_SYSTEME_PC_SNCF_PA_Liaison_PC______PA;
GVL_PIRATE_Interne.E_PLOUIGNEAU_SA_Manque_SA := GVL_PIRATE.PLOUIGNEAU_SA_Manque_SA;
GVL_PIRATE_Interne.E_PLOUIGNEAU_IL2_Inter__de_ligne_2x25kv_V2 := GVL_PIRATE.PLOUIGNEAU_IL2_Inter__de_ligne_2x25kv_V2;
GVL_PIRATE_Interne.E_PLOUIGNEAU_SYSTEME_PA_SNCF_PA_Carte_s__TC := GVL_PIRATE.PLOUIGNEAU_SYSTEME_PA_SNCF_PA_Carte_s__TC;
GVL_PIRATE_Interne.E_PLOUIGNEAU_S4_12_Sect__de_pontage_V2 := GVL_PIRATE.PLOUIGNEAU_S4_12_Sect__de_pontage_V2;
GVL_PIRATE_Interne.E_PLOUIGNEAU_SAT1___25kV_Sect__alimentation_auto_transfo1 := GVL_PIRATE.PLOUIGNEAU_SAT1___25kV_Sect__alimentation_auto_transfo1;
GVL_PIRATE_Interne.E_PLOUIGNEAU_IL4_Inter__de_ligne_2x25kv_V2 := GVL_PIRATE.PLOUIGNEAU_IL4_Inter__de_ligne_2x25kv_V2;
GVL_PIRATE_Interne.E_PLOUIGNEAU_SYSTEME_PC_SNCF_PA_Douteux_vu_du_PC := GVL_PIRATE.PLOUIGNEAU_SYSTEME_PC_SNCF_PA_Douteux_vu_du_PC;
GVL_PIRATE_Interne.E_PLOUIGNEAU_SYSTEME_PC_SNCF_PA_Non_date := GVL_PIRATE.PLOUIGNEAU_SYSTEME_PC_SNCF_PA_Non_date;
GVL_PIRATE_Interne.E_PLOUIGNEAU_SAT2___25kV_Sect__alimentation_auto_transfo2 := GVL_PIRATE.PLOUIGNEAU_SAT2___25kV_Sect__alimentation_auto_transfo2;
GVL_PIRATE_Interne.E_PLOUIGNEAU_SYSTEME_PA_SNCF_PA_Perte_Date := GVL_PIRATE.PLOUIGNEAU_SYSTEME_PA_SNCF_PA_Perte_Date;
GVL_PIRATE_Interne.E_PLOUIGNEAU_IL1_Inter__de_ligne_25kv_V1 := GVL_PIRATE.PLOUIGNEAU_IL1_Inter__de_ligne_25kv_V1;
GVL_PIRATE_Interne.E_PLOUIGNEAU_S5_11_Sect__de_pontage_V1 := GVL_PIRATE.PLOUIGNEAU_S5_11_Sect__de_pontage_V1;
GVL_PIRATE_Interne.E_PLOUIGNEAU_SYSTEME_PC_SNCF_PA_Titulaire := GVL_PIRATE.PLOUIGNEAU_SYSTEME_PC_SNCF_PA_Titulaire;
GVL_PIRATE_Interne.E_PLOUIGNEAU_Contrile_Local_Commande_locale_individuelle := GVL_PIRATE.PLOUIGNEAU_Contrile_Local_Commande_locale_individuelle;
GVL_PIRATE_Interne.E_PLOUIGNEAU_SYSTEME_PA_SNCF_PA_Perte_Information := GVL_PIRATE.PLOUIGNEAU_SYSTEME_PA_SNCF_PA_Perte_Information;
GVL_PIRATE_Interne.E_PLOUIGNEAU_FICTIF_Organe_Fictif := GVL_PIRATE.PLOUIGNEAU_FICTIF_Organe_Fictif;
GVL_PIRATE_Interne.E_PLOUNERIN_IL4_Inter__de_ligne_2x25kv_V2 := GVL_PIRATE.PLOUNERIN_IL4_Inter__de_ligne_2x25kv_V2;
GVL_PIRATE_Interne.E_PLOUNERIN_IL3_Inter__de_ligne_25kv_V1 := GVL_PIRATE.PLOUNERIN_IL3_Inter__de_ligne_25kv_V1;
GVL_PIRATE_Interne.E_PLOUNERIN_SAT2___25kV_Sect__alimentation_auto_transfo2 := GVL_PIRATE.PLOUNERIN_SAT2___25kV_Sect__alimentation_auto_transfo2;
GVL_PIRATE_Interne.E_PLOUNERIN_FICTIF_Organe_Fictif := GVL_PIRATE.PLOUNERIN_FICTIF_Organe_Fictif;
LireEntrees := TRUE;
END_FUNCTION

(* ---- FB_BFS.st ---- *)
FUNCTION_BLOCK FB_BFS
VAR_INPUT
    NbNoeuds : UINT;
    NbAretes : UINT;
    NbEquipements : UINT;
    Sources : ARRAY[0..56] OF BOOL;
    Aretes : ARRAY[0..79] OF ST_AreteZone;
    Equipements : ARRAY[0..79] OF ST_Equipement;
END_VAR
VAR_IN_OUT
    Noeuds : ARRAY[0..56] OF ST_Noeud;
END_VAR
VAR_OUTPUT
    ErreurConfiguration : BOOL;
END_VAR
VAR
    FileNoeuds : ARRAY[0..56] OF UINT;
    TeteFile : UINT;
    FinFile : UINT;
    NoeudCourant : UINT;
    NoeudVoisin : UINT;
    i : INT;
    j : INT;
    k : INT;
    IndexEquipement : INT;
    AreteActive : BOOL;
END_VAR

// Validation des dimensions AVANT toute propagation.
ErreurConfiguration := (NbNoeuds > 57) OR (NbAretes > 80)
    OR (NbEquipements > 80);

IF NOT ErreurConfiguration THEN
    // Verification structurelle : pas d'indices invalides.
    FOR j := 0 TO UINT_TO_INT(NbAretes) - 1 DO
        IndexEquipement := Aretes[j].EquipementIndex;
        IF (Aretes[j].NoeudA >= NbNoeuds)
            OR (Aretes[j].NoeudB >= NbNoeuds)
            OR (IndexEquipement < -1)
            OR (IndexEquipement >= UINT_TO_INT(NbEquipements)) THEN
            ErreurConfiguration := TRUE;
        END_IF;
    END_FOR;
END_IF;

// Un graphe invalide ne doit jamais exposer un etat SousTension obsolete.
FOR i := 0 TO 56 DO
    Noeuds[i].SousTension := FALSE;
END_FOR;

IF NOT ErreurConfiguration THEN
    TeteFile := 0;
    FinFile := 0;

    FOR i := 0 TO UINT_TO_INT(NbNoeuds) - 1 DO
        IF Sources[i] THEN
            Noeuds[i].SousTension := TRUE;
            FileNoeuds[FinFile] := INT_TO_UINT(i);
            FinFile := FinFile + 1;
        END_IF;
    END_FOR;

    WHILE TeteFile < FinFile DO
        NoeudCourant := FileNoeuds[TeteFile];
        TeteFile := TeteFile + 1;

        FOR k := 0 TO UINT_TO_INT(NbAretes) - 1 DO
            IndexEquipement := Aretes[k].EquipementIndex;
            AreteActive := IndexEquipement = -1;
            IF IndexEquipement >= 0 THEN
                AreteActive := Equipements[IndexEquipement].Ferme
                    AND NOT Equipements[IndexEquipement].Defaut;
            END_IF;

            IF AreteActive THEN
                IF Aretes[k].NoeudA = NoeudCourant THEN
                    NoeudVoisin := Aretes[k].NoeudB;
                ELSIF Aretes[k].NoeudB = NoeudCourant THEN
                    NoeudVoisin := Aretes[k].NoeudA;
                ELSE
                    CONTINUE;
                END_IF;

                IF NOT Noeuds[NoeudVoisin].SousTension THEN
                    // Au plus un enfilement par noeud : capacite 57.
                    Noeuds[NoeudVoisin].SousTension := TRUE;
                    FileNoeuds[FinFile] := NoeudVoisin;
                    FinFile := FinFile + 1;
                END_IF;
            END_IF;
        END_FOR;
    END_WHILE;
END_IF;

END_FUNCTION_BLOCK

(* ---- FB_InterfacePIRATE.st ---- *)
FUNCTION_BLOCK FB_InterfacePIRATE
VAR
    // Squelette d'adaptation des variables de supervision.
    // Mapping et polarites non verifies : aucune liaison active.
END_VAR

END_FUNCTION_BLOCK

(* ---- FB_Zone.st ---- *)
FUNCTION_BLOCK FB_Zone
VAR_INPUT
    SourceS11Active : BOOL; // Source Pencran, noeud metier 56
    SourceS21Active : BOOL; // Source Pencran, noeud metier 57
END_VAR
VAR_OUTPUT
    ErreurConfiguration : BOOL;
END_VAR
VAR
    // Coeur du simulateur. Toutes les donnees appartiennent a la zone.
    // Indices 0..56 et 0..79, numérotation metier = indice + 1.
    Noeuds : ARRAY[0..56] OF ST_Noeud;
    Equipements : ARRAY[0..79] OF ST_Equipement;
    Aretes : ARRAY[0..79] OF ST_AreteZone;
    Sources : ARRAY[0..56] OF BOOL;
    NbNoeuds : UINT := 57;
    NbEquipements : UINT := 80;
    NbAretes : UINT := 80;
    ConfigurationChargee : BOOL := FALSE;
    MoteurBFS : FB_BFS;
    i : INT;
END_VAR

// Les 80 equipements sont initialises uniquement au premier cycle.
// En exploitation, definir Equipements[index].Ferme et .Defaut depuis
// l'IHM ou un mapping PIRATE valide, avant l'appel cyclique au FB.
IF NOT ConfigurationChargee THEN
    FOR i := 0 TO 56 DO
        Noeuds[i].IdZone := INT_TO_UINT(i + 1);
        Noeuds[i].SousTension := FALSE;
        Sources[i] := FALSE;
    END_FOR;
    // [0] BREST_IL1 : noeuds 49 - 47
    Equipements[0].Id := 1;
    Equipements[0].Ferme := FALSE;
    Equipements[0].Defaut := FALSE;
    Equipements[0].Asservi := FALSE;
    Equipements[0].Conducteur := FALSE;
    Aretes[0].NoeudA := 48;
    Aretes[0].NoeudB := 46;
    Aretes[0].EquipementIndex := 0;
    // [1] BREST_IL2 : noeuds 49 - 48
    Equipements[1].Id := 2;
    Equipements[1].Ferme := FALSE;
    Equipements[1].Defaut := FALSE;
    Equipements[1].Asservi := FALSE;
    Equipements[1].Conducteur := FALSE;
    Aretes[1].NoeudA := 48;
    Aretes[1].NoeudB := 47;
    Aretes[1].EquipementIndex := 1;
    // [2] KERIVIN_IL1 : noeuds 19 - 13
    Equipements[2].Id := 3;
    Equipements[2].Ferme := FALSE;
    Equipements[2].Defaut := FALSE;
    Equipements[2].Asservi := FALSE;
    Equipements[2].Conducteur := FALSE;
    Aretes[2].NoeudA := 18;
    Aretes[2].NoeudB := 12;
    Aretes[2].EquipementIndex := 2;
    // [3] KERIVIN_IL2 : noeuds 18 - 16
    Equipements[3].Id := 4;
    Equipements[3].Ferme := FALSE;
    Equipements[3].Defaut := FALSE;
    Equipements[3].Asservi := FALSE;
    Equipements[3].Conducteur := FALSE;
    Aretes[3].NoeudA := 17;
    Aretes[3].NoeudB := 15;
    Aretes[3].EquipementIndex := 3;
    // [4] KERIVIN_IL3 : noeuds 19 - 21
    Equipements[4].Id := 5;
    Equipements[4].Ferme := FALSE;
    Equipements[4].Defaut := FALSE;
    Equipements[4].Asservi := FALSE;
    Equipements[4].Conducteur := FALSE;
    Aretes[4].NoeudA := 18;
    Aretes[4].NoeudB := 20;
    Aretes[4].EquipementIndex := 4;
    // [5] KERIVIN_IL4 : noeuds 18 - 22
    Equipements[5].Id := 6;
    Equipements[5].Ferme := FALSE;
    Equipements[5].Defaut := FALSE;
    Equipements[5].Asservi := FALSE;
    Equipements[5].Conducteur := FALSE;
    Aretes[5].NoeudA := 17;
    Aretes[5].NoeudB := 21;
    Aretes[5].EquipementIndex := 5;
    // [6] KERIVIN_IMP : noeuds 18 - 19
    Equipements[6].Id := 7;
    Equipements[6].Ferme := FALSE;
    Equipements[6].Defaut := FALSE;
    Equipements[6].Asservi := FALSE;
    Equipements[6].Conducteur := FALSE;
    Aretes[6].NoeudA := 17;
    Aretes[6].NoeudB := 18;
    Aretes[6].EquipementIndex := 6;
    // [7] KERIVIN_S13-21 : noeuds 13 - 21
    Equipements[7].Id := 8;
    Equipements[7].Ferme := FALSE;
    Equipements[7].Defaut := FALSE;
    Equipements[7].Asservi := FALSE;
    Equipements[7].Conducteur := FALSE;
    Aretes[7].NoeudA := 12;
    Aretes[7].NoeudB := 20;
    Aretes[7].EquipementIndex := 7;
    // [8] KERIVIN_S18-20 : noeuds 16 - 22
    Equipements[8].Id := 9;
    Equipements[8].Ferme := FALSE;
    Equipements[8].Defaut := FALSE;
    Equipements[8].Asservi := FALSE;
    Equipements[8].Conducteur := FALSE;
    Aretes[8].NoeudA := 15;
    Aretes[8].NoeudB := 21;
    Aretes[8].EquipementIndex := 8;
    // [9] KERIVIN_SAT1 : noeuds 19 - 20
    Equipements[9].Id := 10;
    Equipements[9].Ferme := FALSE;
    Equipements[9].Defaut := FALSE;
    Equipements[9].Asservi := FALSE;
    Equipements[9].Conducteur := FALSE;
    Aretes[9].NoeudA := 18;
    Aretes[9].NoeudB := 19;
    Aretes[9].EquipementIndex := 9;
    // [10] KERIVIN_SAT2 : noeuds 17 - 18
    Equipements[10].Id := 11;
    Equipements[10].Ferme := FALSE;
    Equipements[10].Defaut := FALSE;
    Equipements[10].Asservi := FALSE;
    Equipements[10].Conducteur := FALSE;
    Aretes[10].NoeudA := 16;
    Aretes[10].NoeudB := 17;
    Aretes[10].EquipementIndex := 10;
    // [11] LANDERNEAU_I3 : noeuds 37 - 39
    Equipements[11].Id := 12;
    Equipements[11].Ferme := FALSE;
    Equipements[11].Defaut := FALSE;
    Equipements[11].Asservi := FALSE;
    Equipements[11].Conducteur := FALSE;
    Aretes[11].NoeudA := 36;
    Aretes[11].NoeudB := 38;
    Aretes[11].EquipementIndex := 11;
    // [12] LANDERNEAU_I4 : noeuds 38 - 40
    Equipements[12].Id := 13;
    Equipements[12].Ferme := FALSE;
    Equipements[12].Defaut := FALSE;
    Equipements[12].Asservi := FALSE;
    Equipements[12].Conducteur := FALSE;
    Aretes[12].NoeudA := 37;
    Aretes[12].NoeudB := 39;
    Aretes[12].EquipementIndex := 12;
    // [13] LANDIVISIAU_IL1 : noeuds 30 - 27
    Equipements[13].Id := 14;
    Equipements[13].Ferme := FALSE;
    Equipements[13].Defaut := FALSE;
    Equipements[13].Asservi := FALSE;
    Equipements[13].Conducteur := FALSE;
    Aretes[13].NoeudA := 29;
    Aretes[13].NoeudB := 26;
    Aretes[13].EquipementIndex := 13;
    // [14] LANDIVISIAU_IL2 : noeuds 31 - 28
    Equipements[14].Id := 15;
    Equipements[14].Ferme := FALSE;
    Equipements[14].Defaut := FALSE;
    Equipements[14].Asservi := FALSE;
    Equipements[14].Conducteur := FALSE;
    Aretes[14].NoeudA := 30;
    Aretes[14].NoeudB := 27;
    Aretes[14].EquipementIndex := 14;
    // [15] LANDIVISIAU_IL3 : noeuds 30 - 33
    Equipements[15].Id := 16;
    Equipements[15].Ferme := FALSE;
    Equipements[15].Defaut := FALSE;
    Equipements[15].Asservi := FALSE;
    Equipements[15].Conducteur := FALSE;
    Aretes[15].NoeudA := 29;
    Aretes[15].NoeudB := 32;
    Aretes[15].EquipementIndex := 15;
    // [16] LANDIVISIAU_IL4 : noeuds 31 - 34
    Equipements[16].Id := 17;
    Equipements[16].Ferme := FALSE;
    Equipements[16].Defaut := FALSE;
    Equipements[16].Asservi := FALSE;
    Equipements[16].Conducteur := FALSE;
    Aretes[16].NoeudA := 30;
    Aretes[16].NoeudB := 33;
    Aretes[16].EquipementIndex := 16;
    // [17] LANDIVISIAU_IMP : noeuds 30 - 31
    Equipements[17].Id := 18;
    Equipements[17].Ferme := FALSE;
    Equipements[17].Defaut := FALSE;
    Equipements[17].Asservi := FALSE;
    Equipements[17].Conducteur := FALSE;
    Aretes[17].NoeudA := 29;
    Aretes[17].NoeudB := 30;
    Aretes[17].EquipementIndex := 17;
    // [18] LANDIVISIAU_S30-40 : noeuds 28 - 34
    Equipements[18].Id := 19;
    Equipements[18].Ferme := FALSE;
    Equipements[18].Defaut := FALSE;
    Equipements[18].Asservi := FALSE;
    Equipements[18].Conducteur := FALSE;
    Aretes[18].NoeudA := 27;
    Aretes[18].NoeudB := 33;
    Aretes[18].EquipementIndex := 18;
    // [19] LANDIVISIAU_S31-41 : noeuds 27 - 33
    Equipements[19].Id := 20;
    Equipements[19].Ferme := FALSE;
    Equipements[19].Defaut := FALSE;
    Equipements[19].Asservi := FALSE;
    Equipements[19].Conducteur := FALSE;
    Aretes[19].NoeudA := 26;
    Aretes[19].NoeudB := 32;
    Aretes[19].EquipementIndex := 19;
    // [20] LANDIVISIAU_SAT1 : noeuds 29 - 30
    Equipements[20].Id := 21;
    Equipements[20].Ferme := FALSE;
    Equipements[20].Defaut := FALSE;
    Equipements[20].Asservi := FALSE;
    Equipements[20].Conducteur := FALSE;
    Aretes[20].NoeudA := 28;
    Aretes[20].NoeudB := 29;
    Aretes[20].EquipementIndex := 20;
    // [21] LANDIVISIAU_SAT2 : noeuds 31 - 32
    Equipements[21].Id := 22;
    Equipements[21].Ferme := FALSE;
    Equipements[21].Defaut := FALSE;
    Equipements[21].Asservi := FALSE;
    Equipements[21].Conducteur := FALSE;
    Aretes[21].NoeudA := 30;
    Aretes[21].NoeudB := 31;
    Aretes[21].EquipementIndex := 21;
    // [22] LA_FOREST_IMP1 : noeuds 41 - 39
    Equipements[22].Id := 23;
    Equipements[22].Ferme := FALSE;
    Equipements[22].Defaut := FALSE;
    Equipements[22].Asservi := FALSE;
    Equipements[22].Conducteur := FALSE;
    Aretes[22].NoeudA := 40;
    Aretes[22].NoeudB := 38;
    Aretes[22].EquipementIndex := 22;
    // [23] LA_FOREST_IMP2 : noeuds 41 - 40
    Equipements[23].Id := 24;
    Equipements[23].Ferme := FALSE;
    Equipements[23].Defaut := FALSE;
    Equipements[23].Asservi := FALSE;
    Equipements[23].Conducteur := FALSE;
    Aretes[23].NoeudA := 40;
    Aretes[23].NoeudB := 39;
    Aretes[23].EquipementIndex := 23;
    // [24] LA_FOREST_SAT : noeuds 41 - 42
    Equipements[24].Id := 25;
    Equipements[24].Ferme := FALSE;
    Equipements[24].Defaut := FALSE;
    Equipements[24].Asservi := FALSE;
    Equipements[24].Conducteur := FALSE;
    Aretes[24].NoeudA := 40;
    Aretes[24].NoeudB := 41;
    Aretes[24].EquipementIndex := 24;
    // [25] MORLAIX_I13 : noeuds 11 - 13
    Equipements[25].Id := 26;
    Equipements[25].Ferme := FALSE;
    Equipements[25].Defaut := FALSE;
    Equipements[25].Asservi := FALSE;
    Equipements[25].Conducteur := FALSE;
    Aretes[25].NoeudA := 10;
    Aretes[25].NoeudB := 12;
    Aretes[25].EquipementIndex := 25;
    // [26] MORLAIX_I14 : noeuds 12 - 14
    Equipements[26].Id := 27;
    Equipements[26].Ferme := FALSE;
    Equipements[26].Defaut := FALSE;
    Equipements[26].Asservi := FALSE;
    Equipements[26].Conducteur := FALSE;
    Aretes[26].NoeudA := 11;
    Aretes[26].NoeudB := 13;
    Aretes[26].EquipementIndex := 26;
    // [27] MORLAIX_I16 : noeuds 14 - 15
    Equipements[27].Id := 28;
    Equipements[27].Ferme := FALSE;
    Equipements[27].Defaut := FALSE;
    Equipements[27].Asservi := FALSE;
    Equipements[27].Conducteur := FALSE;
    Aretes[27].NoeudA := 13;
    Aretes[27].NoeudB := 14;
    Aretes[27].EquipementIndex := 27;
    // [28] MORLAIX_I18 : noeuds 15 - 16
    Equipements[28].Id := 29;
    Equipements[28].Ferme := FALSE;
    Equipements[28].Defaut := FALSE;
    Equipements[28].Asservi := FALSE;
    Equipements[28].Conducteur := FALSE;
    Aretes[28].NoeudA := 14;
    Aretes[28].NoeudB := 15;
    Aretes[28].EquipementIndex := 28;
    // [29] PENCRAN_D1 : noeuds 50 - 51
    Equipements[29].Id := 30;
    Equipements[29].Ferme := FALSE;
    Equipements[29].Defaut := FALSE;
    Equipements[29].Asservi := FALSE;
    Equipements[29].Conducteur := FALSE;
    Aretes[29].NoeudA := 49;
    Aretes[29].NoeudB := 50;
    Aretes[29].EquipementIndex := 29;
    // [30] PENCRAN_D2 : noeuds 53 - 54
    Equipements[30].Id := 31;
    Equipements[30].Ferme := FALSE;
    Equipements[30].Defaut := FALSE;
    Equipements[30].Asservi := FALSE;
    Equipements[30].Conducteur := FALSE;
    Aretes[30].NoeudA := 52;
    Aretes[30].NoeudB := 53;
    Aretes[30].EquipementIndex := 30;
    // [31] PENCRAN_DB : noeuds 55 - 36
    Equipements[31].Id := 32;
    Equipements[31].Ferme := FALSE;
    Equipements[31].Defaut := FALSE;
    Equipements[31].Asservi := FALSE;
    Equipements[31].Conducteur := FALSE;
    Aretes[31].NoeudA := 54;
    Aretes[31].NoeudB := 35;
    Aretes[31].EquipementIndex := 31;
    // [32] PENCRAN_DL : noeuds 52 - 35
    Equipements[32].Id := 33;
    Equipements[32].Ferme := FALSE;
    Equipements[32].Defaut := FALSE;
    Equipements[32].Asservi := FALSE;
    Equipements[32].Conducteur := FALSE;
    Aretes[32].NoeudA := 51;
    Aretes[32].NoeudB := 34;
    Aretes[32].EquipementIndex := 32;
    // [33] PENCRAN_IS1 : noeuds 35 - 33
    Equipements[33].Id := 34;
    Equipements[33].Ferme := FALSE;
    Equipements[33].Defaut := FALSE;
    Equipements[33].Asservi := FALSE;
    Equipements[33].Conducteur := FALSE;
    Aretes[33].NoeudA := 34;
    Aretes[33].NoeudB := 32;
    Aretes[33].EquipementIndex := 33;
    // [34] PENCRAN_IS2 : noeuds 35 - 34
    Equipements[34].Id := 35;
    Equipements[34].Ferme := FALSE;
    Equipements[34].Defaut := FALSE;
    Equipements[34].Asservi := FALSE;
    Equipements[34].Conducteur := FALSE;
    Aretes[34].NoeudA := 34;
    Aretes[34].NoeudB := 33;
    Aretes[34].EquipementIndex := 34;
    // [35] PENCRAN_IS3 : noeuds 36 - 37
    Equipements[35].Id := 36;
    Equipements[35].Ferme := FALSE;
    Equipements[35].Defaut := FALSE;
    Equipements[35].Asservi := FALSE;
    Equipements[35].Conducteur := FALSE;
    Aretes[35].NoeudA := 35;
    Aretes[35].NoeudB := 36;
    Aretes[35].EquipementIndex := 35;
    // [36] PENCRAN_IS4 : noeuds 36 - 38
    Equipements[36].Id := 37;
    Equipements[36].Ferme := FALSE;
    Equipements[36].Defaut := FALSE;
    Equipements[36].Asservi := FALSE;
    Equipements[36].Conducteur := FALSE;
    Aretes[36].NoeudA := 35;
    Aretes[36].NoeudB := 37;
    Aretes[36].EquipementIndex := 36;
    // [37] PENCRAN_P1 : noeuds 33 - 37
    Equipements[37].Id := 38;
    Equipements[37].Ferme := FALSE;
    Equipements[37].Defaut := FALSE;
    Equipements[37].Asservi := FALSE;
    Equipements[37].Conducteur := FALSE;
    Aretes[37].NoeudA := 32;
    Aretes[37].NoeudB := 36;
    Aretes[37].EquipementIndex := 37;
    // [38] PENCRAN_P2 : noeuds 34 - 38
    Equipements[38].Id := 39;
    Equipements[38].Ferme := FALSE;
    Equipements[38].Defaut := FALSE;
    Equipements[38].Asservi := FALSE;
    Equipements[38].Conducteur := FALSE;
    Aretes[38].NoeudA := 33;
    Aretes[38].NoeudB := 37;
    Aretes[38].EquipementIndex := 38;
    // [39] PENCRAN_S11 : noeuds 56 - 50
    Equipements[39].Id := 40;
    Equipements[39].Ferme := FALSE;
    Equipements[39].Defaut := FALSE;
    Equipements[39].Asservi := FALSE;
    Equipements[39].Conducteur := FALSE;
    Aretes[39].NoeudA := 55;
    Aretes[39].NoeudB := 49;
    Aretes[39].EquipementIndex := 39;
    // [40] PENCRAN_S21 : noeuds 57 - 53
    Equipements[40].Id := 41;
    Equipements[40].Ferme := FALSE;
    Equipements[40].Defaut := FALSE;
    Equipements[40].Asservi := FALSE;
    Equipements[40].Conducteur := FALSE;
    Aretes[40].NoeudA := 56;
    Aretes[40].NoeudB := 52;
    Aretes[40].EquipementIndex := 40;
    // [41] PENCRAN_SB1 : noeuds 52 - 55
    Equipements[41].Id := 42;
    Equipements[41].Ferme := FALSE;
    Equipements[41].Defaut := FALSE;
    Equipements[41].Asservi := FALSE;
    Equipements[41].Conducteur := FALSE;
    Aretes[41].NoeudA := 51;
    Aretes[41].NoeudB := 54;
    Aretes[41].EquipementIndex := 41;
    // [42] PENCRAN_SBP1 : noeuds 50 - 53
    Equipements[42].Id := 43;
    Equipements[42].Ferme := FALSE;
    Equipements[42].Defaut := FALSE;
    Equipements[42].Asservi := FALSE;
    Equipements[42].Conducteur := FALSE;
    Aretes[42].NoeudA := 49;
    Aretes[42].NoeudB := 52;
    Aretes[42].EquipementIndex := 42;
    // [43] PENCRAN_SLB1 : noeuds 35 - 36
    Equipements[43].Id := 44;
    Equipements[43].Ferme := FALSE;
    Equipements[43].Defaut := FALSE;
    Equipements[43].Asservi := FALSE;
    Equipements[43].Conducteur := FALSE;
    Aretes[43].NoeudA := 34;
    Aretes[43].NoeudB := 35;
    Aretes[43].EquipementIndex := 43;
    // [44] PENCRAN_SRB1 : noeuds 51 - 52
    Equipements[44].Id := 45;
    Equipements[44].Ferme := FALSE;
    Equipements[44].Defaut := FALSE;
    Equipements[44].Asservi := FALSE;
    Equipements[44].Conducteur := FALSE;
    Aretes[44].NoeudA := 50;
    Aretes[44].NoeudB := 51;
    Aretes[44].EquipementIndex := 44;
    // [45] PENCRAN_SRB2 : noeuds 54 - 55
    Equipements[45].Id := 46;
    Equipements[45].Ferme := FALSE;
    Equipements[45].Defaut := FALSE;
    Equipements[45].Asservi := FALSE;
    Equipements[45].Conducteur := FALSE;
    Aretes[45].NoeudA := 53;
    Aretes[45].NoeudB := 54;
    Aretes[45].EquipementIndex := 45;
    // [46] PLOUIGNEAU_IL1 : noeuds 9 - 5
    Equipements[46].Id := 47;
    Equipements[46].Ferme := FALSE;
    Equipements[46].Defaut := FALSE;
    Equipements[46].Asservi := FALSE;
    Equipements[46].Conducteur := FALSE;
    Aretes[46].NoeudA := 8;
    Aretes[46].NoeudB := 4;
    Aretes[46].EquipementIndex := 46;
    // [47] PLOUIGNEAU_IL2 : noeuds 8 - 6
    Equipements[47].Id := 48;
    Equipements[47].Ferme := FALSE;
    Equipements[47].Defaut := FALSE;
    Equipements[47].Asservi := FALSE;
    Equipements[47].Conducteur := FALSE;
    Aretes[47].NoeudA := 7;
    Aretes[47].NoeudB := 5;
    Aretes[47].EquipementIndex := 47;
    // [48] PLOUIGNEAU_IL3 : noeuds 9 - 11
    Equipements[48].Id := 49;
    Equipements[48].Ferme := FALSE;
    Equipements[48].Defaut := FALSE;
    Equipements[48].Asservi := FALSE;
    Equipements[48].Conducteur := FALSE;
    Aretes[48].NoeudA := 8;
    Aretes[48].NoeudB := 10;
    Aretes[48].EquipementIndex := 48;
    // [49] PLOUIGNEAU_IL4 : noeuds 8 - 12
    Equipements[49].Id := 50;
    Equipements[49].Ferme := FALSE;
    Equipements[49].Defaut := FALSE;
    Equipements[49].Asservi := FALSE;
    Equipements[49].Conducteur := FALSE;
    Aretes[49].NoeudA := 7;
    Aretes[49].NoeudB := 11;
    Aretes[49].EquipementIndex := 49;
    // [50] PLOUIGNEAU_IMP : noeuds 8 - 9
    Equipements[50].Id := 51;
    Equipements[50].Ferme := FALSE;
    Equipements[50].Defaut := FALSE;
    Equipements[50].Asservi := FALSE;
    Equipements[50].Conducteur := FALSE;
    Aretes[50].NoeudA := 7;
    Aretes[50].NoeudB := 8;
    Aretes[50].EquipementIndex := 50;
    // [51] PLOUIGNEAU_S4-12 : noeuds 6 - 12
    Equipements[51].Id := 52;
    Equipements[51].Ferme := FALSE;
    Equipements[51].Defaut := FALSE;
    Equipements[51].Asservi := FALSE;
    Equipements[51].Conducteur := FALSE;
    Aretes[51].NoeudA := 5;
    Aretes[51].NoeudB := 11;
    Aretes[51].EquipementIndex := 51;
    // [52] PLOUIGNEAU_S5-11 : noeuds 5 - 11
    Equipements[52].Id := 53;
    Equipements[52].Ferme := FALSE;
    Equipements[52].Defaut := FALSE;
    Equipements[52].Asservi := FALSE;
    Equipements[52].Conducteur := FALSE;
    Aretes[52].NoeudA := 4;
    Aretes[52].NoeudB := 10;
    Aretes[52].EquipementIndex := 52;
    // [53] PLOUIGNEAU_SAT1 : noeuds 9 - 10
    Equipements[53].Id := 54;
    Equipements[53].Ferme := FALSE;
    Equipements[53].Defaut := FALSE;
    Equipements[53].Asservi := FALSE;
    Equipements[53].Conducteur := FALSE;
    Aretes[53].NoeudA := 8;
    Aretes[53].NoeudB := 9;
    Aretes[53].EquipementIndex := 53;
    // [54] PLOUIGNEAU_SAT2 : noeuds 7 - 8
    Equipements[54].Id := 55;
    Equipements[54].Ferme := FALSE;
    Equipements[54].Defaut := FALSE;
    Equipements[54].Asservi := FALSE;
    Equipements[54].Conducteur := FALSE;
    Aretes[54].NoeudA := 6;
    Aretes[54].NoeudB := 7;
    Aretes[54].EquipementIndex := 54;
    // [55] PLOUNERIN_IL1 : noeuds 2 - 5
    Equipements[55].Id := 56;
    Equipements[55].Ferme := FALSE;
    Equipements[55].Defaut := FALSE;
    Equipements[55].Asservi := FALSE;
    Equipements[55].Conducteur := FALSE;
    Aretes[55].NoeudA := 1;
    Aretes[55].NoeudB := 4;
    Aretes[55].EquipementIndex := 55;
    // [56] PLOUNERIN_IL2 : noeuds 2 - 6
    Equipements[56].Id := 57;
    Equipements[56].Ferme := FALSE;
    Equipements[56].Defaut := FALSE;
    Equipements[56].Asservi := FALSE;
    Equipements[56].Conducteur := FALSE;
    Aretes[56].NoeudA := 1;
    Aretes[56].NoeudB := 5;
    Aretes[56].EquipementIndex := 56;
    // [57] PLOUNERIN_IL3 : noeuds 3 - 5
    Equipements[57].Id := 58;
    Equipements[57].Ferme := FALSE;
    Equipements[57].Defaut := FALSE;
    Equipements[57].Asservi := FALSE;
    Equipements[57].Conducteur := FALSE;
    Aretes[57].NoeudA := 2;
    Aretes[57].NoeudB := 4;
    Aretes[57].EquipementIndex := 57;
    // [58] PLOUNERIN_IL4 : noeuds 3 - 6
    Equipements[58].Id := 59;
    Equipements[58].Ferme := FALSE;
    Equipements[58].Defaut := FALSE;
    Equipements[58].Asservi := FALSE;
    Equipements[58].Conducteur := FALSE;
    Aretes[58].NoeudA := 2;
    Aretes[58].NoeudB := 5;
    Aretes[58].EquipementIndex := 58;
    // [59] PLOUNERIN_IP : noeuds 2 - 3
    Equipements[59].Id := 60;
    Equipements[59].Ferme := FALSE;
    Equipements[59].Defaut := FALSE;
    Equipements[59].Asservi := FALSE;
    Equipements[59].Conducteur := FALSE;
    Aretes[59].NoeudA := 1;
    Aretes[59].NoeudB := 2;
    Aretes[59].EquipementIndex := 59;
    // [60] PLOUNERIN_SAT1 : noeuds 1 - 2
    Equipements[60].Id := 61;
    Equipements[60].Ferme := FALSE;
    Equipements[60].Defaut := FALSE;
    Equipements[60].Asservi := FALSE;
    Equipements[60].Conducteur := FALSE;
    Aretes[60].NoeudA := 0;
    Aretes[60].NoeudB := 1;
    Aretes[60].EquipementIndex := 60;
    // [61] PLOUNERIN_SAT2 : noeuds 3 - 4
    Equipements[61].Id := 62;
    Equipements[61].Ferme := FALSE;
    Equipements[61].Defaut := FALSE;
    Equipements[61].Asservi := FALSE;
    Equipements[61].Conducteur := FALSE;
    Aretes[61].NoeudA := 2;
    Aretes[61].NoeudB := 3;
    Aretes[61].EquipementIndex := 61;
    // [62] ST_MARC_IL1 : noeuds 44 - 39
    Equipements[62].Id := 63;
    Equipements[62].Ferme := FALSE;
    Equipements[62].Defaut := FALSE;
    Equipements[62].Asservi := FALSE;
    Equipements[62].Conducteur := FALSE;
    Aretes[62].NoeudA := 43;
    Aretes[62].NoeudB := 38;
    Aretes[62].EquipementIndex := 62;
    // [63] ST_MARC_IL2 : noeuds 45 - 40
    Equipements[63].Id := 64;
    Equipements[63].Ferme := FALSE;
    Equipements[63].Defaut := FALSE;
    Equipements[63].Asservi := FALSE;
    Equipements[63].Conducteur := FALSE;
    Aretes[63].NoeudA := 44;
    Aretes[63].NoeudB := 39;
    Aretes[63].EquipementIndex := 63;
    // [64] ST_MARC_IL3 : noeuds 44 - 47
    Equipements[64].Id := 65;
    Equipements[64].Ferme := FALSE;
    Equipements[64].Defaut := FALSE;
    Equipements[64].Asservi := FALSE;
    Equipements[64].Conducteur := FALSE;
    Aretes[64].NoeudA := 43;
    Aretes[64].NoeudB := 46;
    Aretes[64].EquipementIndex := 64;
    // [65] ST_MARC_IL4 : noeuds 45 - 48
    Equipements[65].Id := 66;
    Equipements[65].Ferme := FALSE;
    Equipements[65].Defaut := FALSE;
    Equipements[65].Asservi := FALSE;
    Equipements[65].Conducteur := FALSE;
    Aretes[65].NoeudA := 44;
    Aretes[65].NoeudB := 47;
    Aretes[65].EquipementIndex := 65;
    // [66] ST_MARC_IMP : noeuds 44 - 45
    Equipements[66].Id := 67;
    Equipements[66].Ferme := FALSE;
    Equipements[66].Defaut := FALSE;
    Equipements[66].Asservi := FALSE;
    Equipements[66].Conducteur := FALSE;
    Aretes[66].NoeudA := 43;
    Aretes[66].NoeudB := 44;
    Aretes[66].EquipementIndex := 66;
    // [67] ST_MARC_S4-10 : noeuds 40 - 48
    Equipements[67].Id := 68;
    Equipements[67].Ferme := FALSE;
    Equipements[67].Defaut := FALSE;
    Equipements[67].Asservi := FALSE;
    Equipements[67].Conducteur := FALSE;
    Aretes[67].NoeudA := 39;
    Aretes[67].NoeudB := 47;
    Aretes[67].EquipementIndex := 67;
    // [68] ST_MARC_S5-11 : noeuds 39 - 47
    Equipements[68].Id := 69;
    Equipements[68].Ferme := FALSE;
    Equipements[68].Defaut := FALSE;
    Equipements[68].Asservi := FALSE;
    Equipements[68].Conducteur := FALSE;
    Aretes[68].NoeudA := 38;
    Aretes[68].NoeudB := 46;
    Aretes[68].EquipementIndex := 68;
    // [69] ST_MARC_SAT1 : noeuds 43 - 44
    Equipements[69].Id := 70;
    Equipements[69].Ferme := FALSE;
    Equipements[69].Defaut := FALSE;
    Equipements[69].Asservi := FALSE;
    Equipements[69].Conducteur := FALSE;
    Aretes[69].NoeudA := 42;
    Aretes[69].NoeudB := 43;
    Aretes[69].EquipementIndex := 69;
    // [70] ST_MARC_SAT2 : noeuds 45 - 46
    Equipements[70].Id := 71;
    Equipements[70].Ferme := FALSE;
    Equipements[70].Defaut := FALSE;
    Equipements[70].Asservi := FALSE;
    Equipements[70].Conducteur := FALSE;
    Aretes[70].NoeudA := 44;
    Aretes[70].NoeudB := 45;
    Aretes[70].EquipementIndex := 70;
    // [71] ST_THEGONNEC_IL1 : noeuds 24 - 21
    Equipements[71].Id := 72;
    Equipements[71].Ferme := FALSE;
    Equipements[71].Defaut := FALSE;
    Equipements[71].Asservi := FALSE;
    Equipements[71].Conducteur := FALSE;
    Aretes[71].NoeudA := 23;
    Aretes[71].NoeudB := 20;
    Aretes[71].EquipementIndex := 71;
    // [72] ST_THEGONNEC_IL2 : noeuds 25 - 22
    Equipements[72].Id := 73;
    Equipements[72].Ferme := FALSE;
    Equipements[72].Defaut := FALSE;
    Equipements[72].Asservi := FALSE;
    Equipements[72].Conducteur := FALSE;
    Aretes[72].NoeudA := 24;
    Aretes[72].NoeudB := 21;
    Aretes[72].EquipementIndex := 72;
    // [73] ST_THEGONNEC_IL3 : noeuds 24 - 27
    Equipements[73].Id := 74;
    Equipements[73].Ferme := FALSE;
    Equipements[73].Defaut := FALSE;
    Equipements[73].Asservi := FALSE;
    Equipements[73].Conducteur := FALSE;
    Aretes[73].NoeudA := 23;
    Aretes[73].NoeudB := 26;
    Aretes[73].EquipementIndex := 73;
    // [74] ST_THEGONNEC_IL4 : noeuds 25 - 28
    Equipements[74].Id := 75;
    Equipements[74].Ferme := FALSE;
    Equipements[74].Defaut := FALSE;
    Equipements[74].Asservi := FALSE;
    Equipements[74].Conducteur := FALSE;
    Aretes[74].NoeudA := 24;
    Aretes[74].NoeudB := 27;
    Aretes[74].EquipementIndex := 74;
    // [75] ST_THEGONNEC_IMP : noeuds 24 - 25
    Equipements[75].Id := 76;
    Equipements[75].Ferme := FALSE;
    Equipements[75].Defaut := FALSE;
    Equipements[75].Asservi := FALSE;
    Equipements[75].Conducteur := FALSE;
    Aretes[75].NoeudA := 23;
    Aretes[75].NoeudB := 24;
    Aretes[75].EquipementIndex := 75;
    // [76] ST_THEGONNEC_S20-30 : noeuds 22 - 28
    Equipements[76].Id := 77;
    Equipements[76].Ferme := FALSE;
    Equipements[76].Defaut := FALSE;
    Equipements[76].Asservi := FALSE;
    Equipements[76].Conducteur := FALSE;
    Aretes[76].NoeudA := 21;
    Aretes[76].NoeudB := 27;
    Aretes[76].EquipementIndex := 76;
    // [77] ST_THEGONNEC_S21-31 : noeuds 21 - 27
    Equipements[77].Id := 78;
    Equipements[77].Ferme := FALSE;
    Equipements[77].Defaut := FALSE;
    Equipements[77].Asservi := FALSE;
    Equipements[77].Conducteur := FALSE;
    Aretes[77].NoeudA := 20;
    Aretes[77].NoeudB := 26;
    Aretes[77].EquipementIndex := 77;
    // [78] ST_THEGONNEC_SAT1 : noeuds 23 - 24
    Equipements[78].Id := 79;
    Equipements[78].Ferme := FALSE;
    Equipements[78].Defaut := FALSE;
    Equipements[78].Asservi := FALSE;
    Equipements[78].Conducteur := FALSE;
    Aretes[78].NoeudA := 22;
    Aretes[78].NoeudB := 23;
    Aretes[78].EquipementIndex := 78;
    // [79] ST_THEGONNEC_SAT2 : noeuds 25 - 26
    Equipements[79].Id := 80;
    Equipements[79].Ferme := FALSE;
    Equipements[79].Defaut := FALSE;
    Equipements[79].Asservi := FALSE;
    Equipements[79].Conducteur := FALSE;
    Aretes[79].NoeudA := 24;
    Aretes[79].NoeudB := 25;
    Aretes[79].EquipementIndex := 79;
    ConfigurationChargee := TRUE;
END_IF;

// Etats derives, pas de valeur Forcee : le defaut coupe sans modifier Ferme.
FOR i := 0 TO 79 DO
    Equipements[i].Conducteur :=
        Equipements[i].Ferme AND NOT Equipements[i].Defaut;
END_FOR;

// Uniquement deux noeuds source, tous les autres restent a FALSE.
Sources[55] := SourceS11Active;
Sources[56] := SourceS21Active;

MoteurBFS(
    NbNoeuds := NbNoeuds,
    NbAretes := NbAretes,
    NbEquipements := NbEquipements,
    Sources := Sources,
    Aretes := Aretes,
    Equipements := Equipements,
    Noeuds := Noeuds
);
ErreurConfiguration := MoteurBFS.ErreurConfiguration;

END_FUNCTION_BLOCK
